TYPE E_CamApplicationError :
(
    CAM_ERROR_NONE := 0,
    CAM_ERROR_COMMAND_NOT_ALLOWED,
    CAM_ERROR_NOT_REFERENCED,
    CAM_ERROR_RECIPE_PITCH,
    CAM_ERROR_RECIPE_CONVEYOR_VELOCITY,
    CAM_ERROR_RECIPE_CUT_VELOCITY,
    CAM_ERROR_RECIPE_EDGE_LENGTH,
    CAM_ERROR_RECIPE_PHASE_ORDER,
    CAM_ERROR_RECIPE_SYNC_SPACE,
    CAM_ERROR_RECIPE_RETURN_SPACE,
    CAM_ERROR_RECIPE_DYNAMICS,
    CAM_ERROR_AXIS_POWER,
    CAM_ERROR_AXIS_REFERENCE,
    CAM_ERROR_CAM_BUILD,
    CAM_ERROR_CAM_LOAD,
    CAM_ERROR_CAM_CHARACTERISTICS,
    CAM_ERROR_CAM_IN,
    CAM_ERROR_MASTER_MOVE,
    CAM_ERROR_MASTER_STOP,
    CAM_ERROR_CAM_OUT,
    CAM_ERROR_SLAVE_RETURN,
    CAM_ERROR_AXIS_RESET
);
END_TYPE

(* stored: Version 1.1.0.1, ProductVersion 3.1.4024.16
   DUT E_CamApplicationError: Id {5be5f029-58e8-401d-8cf9-7b4cc8d4d40c} *)
